FUNCTION_BLOCK FB_HardwareInputs
VAR_OUTPUT
    stInputs : ST_HomeInputs;
END_VAR


stInputs.Workshop.bButton := GVL_WorkshopIO.bButton;
stInputs.Entryway.bLowerButton := GVL_EntrywayIO.bLowerButton;
stInputs.Entryway.bUpperButton := GVL_EntrywayIO.bUpperButton;
stInputs.Hall.bUpperButton := GVL_HallIO.bUpperButton;
stInputs.Hall.bLowerButton := GVL_HallIO.bLowerButton;

END_FUNCTION_BLOCK

(* stored: Version 1.1.0.1
   POU FB_HardwareInputs: Id {c0797200-451f-46aa-8a44-cd6f33cc8863}, SpecialFunc None *)
